(* Production-style program with a FB_KBO_Coating_States nested in FB_KBOInitHost. It follows
   PRG_ATMInit: one motor, the PMPS state-name configurators and the host. The
   arbiter, fast-fault output, persistent storage and DB reader are shared in
   GVL_PRG and ticked by PRG_PMPS_PRE and PRG_PMPS_POST. The configurators are in
   the PRG, because the host's references are not bound yet when its
   declaration initialisers run. The PMPS DB is plc-cc-motion.json. *)
PROGRAM PRG_KBO
VAR
    {attribute 'TcNcAxis' := 'PRG_KBO_Y'}
    axRef         : AXIS_REF;
    fbMotor       : FB_MotionStageNC(
        AxisRef                := axRef,
        iPersistentDataStorage := GVL_PRG.fbPDS,
        sName                  := 'KBOINIT'
    );
    aiMotionStage : ARRAY[1..MotionConstants.MAX_STATE_MOTORS] OF I_MotionStage := [fbMotor];

    astPositionState : ARRAY[1..MotionConstants.MAX_STATE_MOTORS]
                         OF ARRAY[1..GeneralConstants.MAX_STATES] OF ST_PositionState;
    stDefault : ST_PositionState := (
        bMoveOk       := TRUE,
        bValid        := TRUE,
        bUseRawCounts := TRUE
    );
    afbStatePMPS : ARRAY[1..2] OF FB_CC_StatePMPSEncConfig[
        (stPositionState := astPositionState[1][E_KBO_CoatingStates.Si],
         stDefault       := stDefault,
         nEncoderCount   := 1000,
         sPmpsState      := 'TST:KBO-Si'),
        (stPositionState := astPositionState[1][E_KBO_CoatingStates.B4C],
         stDefault       := stDefault,
         nEncoderCount   := 2000,
         sPmpsState      := 'TST:KBO-B4C')
    ];

    fbHost : FB_KBOHost(
        aiMotionStage         := aiMotionStage,
        astPositionState      := astPositionState,
        fbFFHWO               := GVL_PRG.fbFastFaultOutput1,
        fbArbiter             := GVL_PRG.fbArbiter1,
        sDeviceName           := 'TST:KBO',
        sTransitionKey        := 'TST:KBO-TRANSITION',
        bEnableBeamParams     := TRUE,
        bEnablePositionLimits := TRUE,
        bReadDBNow            := TRUE,
        bFileReaderBusy       := MOTION_GVL.fbPmpsFileReader.bBusy,
        bFileReaderError      := MOTION_GVL.fbPmpsFileReader.bError
    );

    i          : UINT;
    bFirstScan : BOOL := TRUE;
END_VAR

IF bFirstScan THEN
    fbMotor.SetModeEnableLimits(
        LimBackward    := TRUE,
        LimForward     := TRUE,
        HomeEnable     := FALSE,
        BrakeMode      := E_StageBrakeMode.IF_ENABLED,
        EnableMode     := E_StageEnableMode.DURING_MOTION,
        HomeMode       := E_EpicsHomeCmd.LOW_LIMIT,
        UserEnable     := TRUE,
        HardwareEnable := TRUE
    );
    fbMotor.SetVelocity(
        Velocity := 15.5
    );
    fbMotor.RestoreMotionParams      := FALSE;
    fbMotor.DoNotRestoreNcParameters := TRUE;
    bFirstScan := FALSE;
END_IF

FOR i := 1 TO 2 DO
    afbStatePMPS[i]();
END_FOR

fbHost();
fbMotor();

END_PROGRAM

(* stored: Version 1.1.0.1
   POU PRG_KBO: Id {bde349c7-37da-44e8-9437-9afa8e527dda}, SpecialFunc None *)
